// TIA Portal V20 export
TYPE "WT2_Kd_Befehl_UDT"
   STRUCT
      iHandshake : Int;
      Befehl : Struct
         iID : Int;
         iParam : Int;
      END_STRUCT;
      Param : Struct
         diID : DInt;
         diValue : DInt;
         iDiv : Int;
         byEditKonfigSet : Byte;
         byReserve : Byte;
         diReserve2 : DInt;
      END_STRUCT;
      FernVorgabeDig : Struct
         bFreigabeNiveaureg : Bool;
         bSollwertumschAB : Bool;
         b222_Reserve : Bool;
         b223_Reserve : Bool;
         b224_Reserve : Bool;
         b225_Reserve : Bool;
         b226_Reserve : Bool;
         b227_Reserve : Bool;
         by23_Reserve : Byte;
      END_STRUCT;
      rFernSollwert : Real;
      byReserve : Array[0..3] of Byte;
   END_STRUCT;
END_TYPE
